(* IEC 61131-3 sources: nautilus/tools/rig/smoke/fixtures/logix-tp, 1 file *)

(* ---- Main.st ---- *)
PROGRAM Main
VAR_EXTERNAL
    Go  : BOOL;
    Out : BOOL;
END_VAR
VAR
    pulse : TP;
END_VAR
pulse(IN := Go, PT := T#500MS);
Out := pulse.Q;
END_PROGRAM
